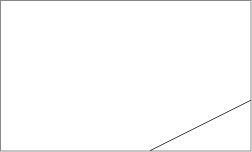
VISUALIZATION VisuC6x  // 252x152
    Line (150,150) (250,100)
END_VISUALIZATION

(* stored: Version 1.1.0.1
   Visu VisuC6x: Id {d69ea30a-a88f-417e-8713-95e2e6cd171c} *)
